      R_g[4,13] := -0.45977530;
      R_g[4,14] := 0.29049909;
      R_g[4,15] := 0.84397930;
      R_g[5,0] := 0.11107527;
      R_g[5,1] := 0.19470578;
      R_g[5,2] := -0.14108169;
      R_g[5,3] := 0.05879988;
      R_g[5,4] := 0.18819207;
      R_g[5,5] := -2.47536159;
      R_g[5,6] := -0.06510852;
      R_g[5,7] := 0.20388806;
      R_g[5,8] := -0.11789436;
      R_g[5,9] := -0.20122005;
      R_g[5,10] := 0.13310707;
      R_g[5,11] := 0.10226060;
      R_g[5,12] := 0.11609720;
      R_g[5,13] := -0.01743704;
      R_g[5,14] := 0.00398547;
      R_g[5,15] := -0.15065657;
      R_g[6,0] := 0.01830370;
      R_g[6,1] := -0.12926060;
      R_g[6,2] := 0.03696303;
      R_g[6,3] := 0.16922043;
      R_g[6,4] := -0.01032830;
      R_g[6,5] := 0.17732817;
      R_g[6,6] := -2.69588876;
      R_g[6,7] := 0.02693873;
      R_g[6,8] := 0.12963313;
      R_g[6,9] := -0.13445157;
      R_g[6,10] := 0.03944382;
      R_g[6,11] := 0.48681569;
      R_g[6,12] := -0.06957243;
      R_g[6,13] := 0.15626159;
      R_g[6,14] := 0.08367650;
      R_g[6,15] := 0.12336652;
      R_g[7,0] := -0.03125253;
      R_g[7,1] := -0.06615835;
      R_g[7,2] := -0.30859804;
      R_g[7,3] := -0.25204793;
      R_g[7,4] := 0.40157086;
      R_g[7,5] := 0.02905789;
      R_g[7,6] := -0.05298730;
      R_g[7,7] := -3.66701341;
      R_g[7,8] := -0.20909342;
      R_g[7,9] := 0.39114916;
      R_g[7,10] := 0.02195679;
      R_g[7,11] := 0.36044669;
      R_g[7,12] := -0.19184318;
      R_g[7,13] := 0.29045779;
      R_g[7,14] := -0.39132181;
      R_g[7,15] := 0.18133201;
      R_g[8,0] := 0.10109203;
      R_g[8,1] := 0.70265359;
      R_g[8,2] := -0.20131305;
      R_g[8,3] := -0.26565599;
      R_g[8,4] := -0.09981477;
      R_g[8,5] := 0.02134162;
      R_g[8,6] := 0.03664974;
      R_g[8,7] := -0.10195713;
      R_g[8,8] := -2.91001201;
      R_g[8,9] := 0.11249696;
      R_g[8,10] := 0.27498955;
      R_g[8,11] := -0.21615753;
      R_g[8,12] := 0.21132010;
      R_g[8,13] := -0.04111291;
      R_g[8,14] := 0.16867815;
      R_g[8,15] := -0.19916441;
      R_g[9,0] := -0.17235202;
      R_g[9,1] := -0.51918679;
      R_g[9,2] := 0.09489006;
      R_g[9,3] := 0.27006283;
      R_g[9,4] := -0.08789669;
      R_g[9,5] := 0.00435399;
      R_g[9,6] := 0.16746791;
      R_g[9,7] := -0.05963518;
      R_g[9,8] := -0.02752298;
      R_g[9,9] := -4.96825457;
      R_g[9,10] := -0.22408967;
      R_g[9,11] := 0.39007574;
      R_g[9,12] := 0.04636907;
      R_g[9,13] := 0.04828465;
      R_g[9,14] := -0.23503923;
      R_g[9,15] := 0.62594104;
      R_g[10,0] := -0.15698923;
      R_g[10,1] := 0.66038901;
      R_g[10,2] := -0.36404622;
      R_g[10,3] := -0.15719211;
      R_g[10,4] := 0.19071013;
      R_g[10,5] := -0.04058476;
      R_g[10,6] := -0.03078617;
      R_g[10,7] := 0.71735823;
      R_g[10,8] := -0.29184514;
      R_g[10,9] := -0.10818060;
      R_g[10,10] := -3.58587956;
      R_g[10,11] := -0.47085500;
      R_g[10,12] := 0.49304882;
      R_g[10,13] := 0.30396828;
      R_g[10,14] := 0.08089786;
      R_g[10,15] := -0.43142110;
      R_g[11,0] := 0.06635704;
      R_g[11,1] := 0.43992752;
      R_g[11,2] := 0.07202107;
      R_g[11,3] := -0.23624249;
      R_g[11,4] := -0.07328893;
      R_g[11,5] := -0.04814436;
      R_g[11,6] := -0.09117863;
      R_g[11,7] := 0.11876864;
      R_g[11,8] := 0.00884132;
      R_g[11,9] := -0.18132856;
      R_g[11,10] := 0.01293289;
      R_g[11,11] := -3.54570603;
      R_g[11,12] := -0.03885806;
      R_g[11,13] := -0.05033415;
      R_g[11,14] := 0.11649126;
      R_g[11,15] := -0.00223985;
      R_g[12,0] := -0.17420630;
      R_g[12,1] := -0.13533008;
      R_g[12,2] := -0.02006780;
      R_g[12,3] := 0.22674133;
      R_g[12,4] := -0.14372772;
      R_g[12,5] := 0.17432602;
      R_g[12,6] := 0.28012389;
      R_g[12,7] := -0.08454837;
      R_g[12,8] := 0.17622249;
      R_g[12,9] := -0.18562099;
      R_g[12,10] := -0.13753660;
      R_g[12,11] := 0.31376547;
      R_g[12,12] := -2.33639669;
      R_g[12,13] := -0.37101883;
      R_g[12,14] := -0.10402304;
      R_g[12,15] := 0.34098265;
      R_g[13,0] := 0.05532536;
      R_g[13,1] := -1.13573086;
      R_g[13,2] := 0.05515465;
      R_g[13,3] := 0.17128730;
      R_g[13,4] := 0.29013124;
      R_g[13,5] := 0.14211339;
      R_g[13,6] := -0.12067565;
      R_g[13,7] := 0.06888673;
      R_g[13,8] := -0.19051172;
      R_g[13,9] := -0.08930715;
      R_g[13,10] := -0.03726633;
      R_g[13,11] := 0.10250945;
      R_g[13,12] := 0.01444966;
      R_g[13,13] := -2.59691453;
      R_g[13,14] := -0.05213837;
      R_g[13,15] := -0.16357523;
      R_g[14,0] := -0.07426858;
      R_g[14,1] := 0.95711172;
      R_g[14,2] := -0.52914786;
      R_g[14,3] := -0.50707346;
      R_g[14,4] := -0.18582524;
      R_g[14,5] := 0.04817829;
      R_g[14,6] := -0.18424018;
      R_g[14,7] := 0.31674099;
      R_g[14,8] := -0.00767360;
      R_g[14,9] := -0.00882705;
      R_g[14,10] := -0.06244185;
      R_g[14,11] := -0.83984315;
      R_g[14,12] := -0.04242671;
      R_g[14,13] := 0.06255507;
      R_g[14,14] := -2.18376112;
      R_g[14,15] := -0.50745595;
      R_g[15,0] := -0.24544616;
      R_g[15,1] := -0.38065434;
      R_g[15,2] := 0.52168375;
      R_g[15,3] := 0.63476181;
      R_g[15,4] := -0.70045185;
      R_g[15,5] := 0.03916581;
      R_g[15,6] := 0.27065009;
      R_g[15,7] := -0.15145577;
      R_g[15,8] := 0.19062088;
      R_g[15,9] := -0.16805187;
      R_g[15,10] := -0.02476993;
      R_g[15,11] := 0.03592181;
      R_g[15,12] := -0.40066659;
      R_g[15,13] := -0.61348122;
      R_g[15,14] := 0.08364772;
      R_g[15,15] := -3.36107063;
      R_o[0,0] := -0.17998135;
      R_o[0,1] := -1.60253966;
      R_o[0,2] := 0.68840933;
      R_o[0,3] := 0.60407180;
      R_o[0,4] := -0.62490994;
      R_o[0,5] := 0.50324053;
      R_o[0,6] := 0.24965659;
      R_o[0,7] := 0.27685815;
      R_o[0,8] := -0.37989971;
      R_o[0,9] := 0.13533561;
      R_o[0,10] := -0.25785661;
      R_o[0,11] := -0.51081169;
      R_o[0,12] := -1.26113296;
      R_o[0,13] := 0.09709056;
      R_o[0,14] := 0.61411685;
      R_o[0,15] := 0.22855295;
      R_o[1,0] := 0.22900739;
      R_o[1,1] := -3.14904022;
      R_o[1,2] := 0.71979213;
      R_o[1,3] := 0.13460559;
      R_o[1,4] := 0.28159738;
      R_o[1,5] := -1.25828946;
      R_o[1,6] := 0.70830607;
      R_o[1,7] := -0.61551344;
      R_o[1,8] := -0.20931304;
      R_o[1,9] := 0.84665543;
      R_o[1,10] := -0.58804363;
      R_o[1,11] := -0.01368906;
      R_o[1,12] := -0.09546302;
      R_o[1,13] := 0.68291515;
      R_o[1,14] := 0.83152312;
      R_o[1,15] := -0.27614936;
      R_o[2,0] := 0.22624512;
      R_o[2,1] := -0.50015140;
      R_o[2,2] := -0.05820123;
      R_o[2,3] := 0.24992104;
      R_o[2,4] := -0.42781389;
      R_o[2,5] := -0.01809851;
      R_o[2,6] := -0.01348706;
      R_o[2,7] := -0.39746183;
      R_o[2,8] := -0.21094593;
      R_o[2,9] := 0.74206448;
      R_o[2,10] := 0.08259194;
      R_o[2,11] := -0.43268228;
      R_o[2,12] := -0.06109180;
      R_o[2,13] := -0.26904088;
      R_o[2,14] := 0.29712129;
      R_o[2,15] := -0.07692748;
      R_o[3,0] := 0.14433832;
      R_o[3,1] := -0.80342203;
      R_o[3,2] := 0.15820050;
      R_o[3,3] := 0.08200698;
      R_o[3,4] := -0.48171204;
      R_o[3,5] := -0.11591465;
      R_o[3,6] := -0.19669321;
      R_o[3,7] := -0.14903167;
      R_o[3,8] := -0.15372486;
      R_o[3,9] := 0.14865009;
      R_o[3,10] := -0.82148689;
      R_o[3,11] := 0.27812725;
      R_o[3,12] := 0.00223510;
      R_o[3,13] := 0.21079217;
      R_o[3,14] := -0.25288963;
      R_o[3,15] := -0.22805665;
      R_o[4,0] := 0.25114408;
      R_o[4,1] := -0.04965499;
      R_o[4,2] := -0.07762759;
      R_o[4,3] := 0.18927185;
      R_o[4,4] := 0.10361283;
      R_o[4,5] := -0.03912014;
      R_o[4,6] := -0.91816306;
      R_o[4,7] := 0.15886311;
      R_o[4,8] := 0.42278275;
      R_o[4,9] := 0.42559728;
      R_o[4,10] := -0.16750900;
      R_o[4,11] := -0.82801008;
      R_o[4,12] := 0.47436076;
      R_o[4,13] := 0.45988649;
      R_o[4,14] := 0.03260082;
      R_o[4,15] := -0.05795699;
      R_o[5,0] := 0.01105135;
      R_o[5,1] := -1.15132201;
      R_o[5,2] := 0.54602605;
      R_o[5,3] := 0.71394539;
      R_o[5,4] := -0.17321546;
      R_o[5,5] := -0.52846497;
      R_o[5,6] := -0.43260244;
      R_o[5,7] := 0.35832340;
      R_o[5,8] := 0.21435645;
      R_o[5,9] := 0.26636124;
      R_o[5,10] := 0.00893501;
      R_o[5,11] := -0.63832158;
      R_o[5,12] := -0.11683670;
      R_o[5,13] := -0.02273753;
      R_o[5,14] := 0.03232908;
      R_o[5,15] := 0.10529289;
      R_o[6,0] := 0.31001085;
      R_o[6,1] := -1.19092143;
      R_o[6,2] := 0.21876206;
      R_o[6,3] := 0.33240157;
      R_o[6,4] := -0.18906151;
      R_o[6,5] := 0.48293993;
      R_o[6,6] := -0.03892522;
      R_o[6,7] := -0.35924369;
      R_o[6,8] := 0.12160594;
      R_o[6,9] := -0.40936342;
      R_o[6,10] := 0.12075932;
      R_o[6,11] := -0.49636525;
      R_o[6,12] := -0.13716739;
      R_o[6,13] := 0.06098676;
      R_o[6,14] := -0.27069107;
      R_o[6,15] := 0.41007137;
      R_o[7,0] := 0.29690558;
      R_o[7,1] := -0.37541282;
      R_o[7,2] := 0.24571100;
      R_o[7,3] := 0.23365253;
      R_o[7,4] := 0.21465455;
      R_o[7,5] := 0.03528690;
      R_o[7,6] := -0.12078243;
      R_o[7,7] := -0.03139850;
      R_o[7,8] := 0.10045099;
      R_o[7,9] := -0.14713535;
      R_o[7,10] := -0.18440804;
      R_o[7,11] := 0.56326222;
      R_o[7,12] := -0.29376999;
      R_o[7,13] := 0.06893768;
      R_o[7,14] := 0.13139424;
      R_o[7,15] := 0.26108429;
      R_o[8,0] := -1.83918154;
      R_o[8,1] := -1.09582520;
      R_o[8,2] := 0.50053239;
      R_o[8,3] := 0.73636478;
      R_o[8,4] := -0.94267857;
      R_o[8,5] := -1.52087641;
      R_o[8,6] := 2.80385971;
      R_o[8,7] := 0.62324148;
      R_o[8,8] := -3.54411769;
      R_o[8,9] := -0.25437289;
      R_o[8,10] := -0.15810332;
      R_o[8,11] := -0.51360112;
      R_o[8,12] := 0.01348928;
      R_o[8,13] := 0.22060399;
      R_o[8,14] := -0.52212816;
      R_o[8,15] := 0.10016742;
      R_o[9,0] := -1.07547414;
      R_o[9,1] := -1.28275371;
      R_o[9,2] := 0.35765028;
      R_o[9,3] := 0.44110700;
      R_o[9,4] := -0.91392058;
      R_o[9,5] := -1.19914532;
      R_o[9,6] := 0.03312799;
      R_o[9,7] := 0.26320797;
      R_o[9,8] := -0.30888504;
      R_o[9,9] := -3.75967288;
      R_o[9,10] := -0.26503733;
      R_o[9,11] := -0.14797226;
      R_o[9,12] := -0.29307473;
      R_o[9,13] := 0.29319406;
      R_o[9,14] := 0.47096246;
      R_o[9,15] := 0.08412670;
      R_o[10,0] := 0.03535339;
      R_o[10,1] := -0.81770265;
      R_o[10,2] := -0.41774553;
      R_o[10,3] := 0.28629521;
      R_o[10,4] := -0.29024190;
      R_o[10,5] := -0.30073890;
      R_o[10,6] := 0.06244223;
      R_o[10,7] := -0.86978775;
      R_o[10,8] := 0.56519794;
      R_o[10,9] := 0.02823679;
      R_o[10,10] := 0.43152261;
      R_o[10,11] := -0.52289534;
      R_o[10,12] := -0.92306936;
      R_o[10,13] := -0.11299136;
      R_o[10,14] := -0.46108496;
      R_o[10,15] := 0.27689543;
      R_o[11,0] := -0.27377477;
      R_o[11,1] := -1.38200986;
      R_o[11,2] := 0.80172545;
      R_o[11,3] := 0.47983712;
      R_o[11,4] := -0.61602306;
      R_o[11,5] := 0.14996068;
      R_o[11,6] := -0.27008256;
      R_o[11,7] := 0.01958398;
      R_o[11,8] := 0.95527297;
      R_o[11,9] := -0.14984407;
      R_o[11,10] := -0.12444744;
      R_o[11,11] := 2.54292870;
      R_o[11,12] := -0.39212865;
      R_o[11,13] := -1.04945409;
      R_o[11,14] := 0.45311722;
      R_o[11,15] := 0.23906973;
      R_o[12,0] := -0.03170222;
      R_o[12,1] := -0.25899503;
      R_o[12,2] := -0.00625280;
      R_o[12,3] := 0.20854484;
      R_o[12,4] := -0.24143498;
      R_o[12,5] := 0.10468624;
      R_o[12,6] := -0.20445421;
      R_o[12,7] := 0.37825984;
      R_o[12,8] := 0.04627231;
      R_o[12,9] := 0.02643433;
      R_o[12,10] := -0.13525262;
      R_o[12,11] := -0.51159739;
      R_o[12,12] := 0.17827436;
      R_o[12,13] := 0.03084075;
      R_o[12,14] := 0.28973144;
      R_o[12,15] := -0.25529897;
      R_o[13,0] := 0.00229840;
      R_o[13,1] := -1.61626279;
      R_o[13,2] := 0.40775979;
      R_o[13,3] := 0.59826922;
      R_o[13,4] := -0.21434167;
      R_o[13,5] := -0.15114538;
      R_o[13,6] := -0.73304671;
      R_o[13,7] := -0.11104193;
      R_o[13,8] := -0.43963873;
      R_o[13,9] := 0.18838404;
      R_o[13,10] := 0.39571330;
      R_o[13,11] := -1.05748773;
      R_o[13,12] := -0.32323301;
      R_o[13,13] := 1.01370287;
      R_o[13,14] := 0.21895173;
      R_o[13,15] := 0.80038011;
      R_o[14,0] := -0.07648548;
      R_o[14,1] := -1.30468404;
      R_o[14,2] := 0.58321625;
      R_o[14,3] := 0.72309285;
      R_o[14,4] := 0.12278607;
      R_o[14,5] := 0.20592272;
      R_o[14,6] := -1.31852913;
      R_o[14,7] := -0.26429388;
      R_o[14,8] := 0.67733824;
      R_o[14,9] := 0.28490099;
      R_o[14,10] := 0.50044572;
      R_o[14,11] := 1.13938892;
      R_o[14,12] := -0.62636727;
      R_o[14,13] := -0.64233524;
      R_o[14,14] := 2.21524429;
      R_o[14,15] := 0.10953581;
      R_o[15,0] := -0.61134338;
      R_o[15,1] := -1.14686418;
      R_o[15,2] := 0.91901773;
      R_o[15,3] := 0.59483540;
      R_o[15,4] := -1.43020630;
      R_o[15,5] := -0.02133927;
      R_o[15,6] := 0.24188809;
      R_o[15,7] := -0.50801885;
      R_o[15,8] := 0.25780970;
      R_o[15,9] := 0.13150303;
      R_o[15,10] := 0.06579445;
      R_o[15,11] := 0.21622118;
      R_o[15,12] := -0.23762867;
      R_o[15,13] := -0.99601251;
      R_o[15,14] := 0.53441352;
      R_o[15,15] := 2.04913473;
      B_i[0] := 2.13055468;
      B_i[1] := -0.28939855;
      B_i[2] := 2.50660825;
      B_i[3] := -0.09900541;
      B_i[4] := 0.92722613;
      B_i[5] := -0.24022682;
      B_i[6] := 0.01314271;
      B_i[7] := -0.16002662;
      B_i[8] := -0.13514934;
      B_i[9] := -0.66461527;
      B_i[10] := -0.39439538;
      B_i[11] := -0.72713459;
      B_i[12] := 2.69549060;
      B_i[13] := 0.10082641;
      B_i[14] := 0.18705003;
      B_i[15] := -0.52215415;
      B_f[0] := 1.71853232;
      B_f[1] := 0.52807707;
      B_f[2] := -0.91032523;
      B_f[3] := -0.51656717;
      B_f[4] := 3.52749252;
      B_f[5] := 2.54868436;
      B_f[6] := 2.06901407;
      B_f[7] := 4.24917698;
      B_f[8] := 2.06338930;
      B_f[9] := 2.86993122;
      B_f[10] := 3.17252159;
      B_f[11] := 1.42340124;
      B_f[12] := 4.81506538;
      B_f[13] := 1.14250445;
      B_f[14] := 0.49386898;
      B_f[15] := 2.75026822;
      B_g[0] := -0.07227773;
      B_g[1] := -0.66488314;
      B_g[2] := 0.70045793;
      B_g[3] := 0.98024452;
      B_g[4] := -0.46857694;
      B_g[5] := 0.02956967;
      B_g[6] := 0.27909416;
      B_g[7] := -0.22752739;
      B_g[8] := -0.10114017;
      B_g[9] := -0.10326473;
      B_g[10] := 0.06763726;
      B_g[11] := 0.14730735;
      B_g[12] := -0.17682402;
      B_g[13] := -0.28040373;
      B_g[14] := 0.69763172;
      B_g[15] := -0.60094702;
      B_o[0] := 3.63638949;
      B_o[1] := 3.95470619;
      B_o[2] := 2.86919069;
      B_o[3] := 2.67019081;
      B_o[4] := 2.45756173;
      B_o[5] := 2.80873203;
      B_o[6] := 2.80962849;
      B_o[7] := 1.47691143;
      B_o[8] := 4.80254173;
      B_o[9] := 3.77295828;
      B_o[10] := 3.93514633;
      B_o[11] := 3.18298674;
      B_o[12] := 1.06958044;
      B_o[13] := 3.72094917;
      B_o[14] := 2.60961676;
      B_o[15] := 3.24567151;
      FC_W[0,0] := -0.82467866;
      FC_W[0,1] := 0.23118977;
      FC_W[0,2] := -0.56444192;
      FC_W[0,3] := -0.32562086;
      FC_W[0,4] := 0.93298566;
      FC_W[0,5] := -1.32120907;
      FC_W[0,6] := -0.26805392;
      FC_W[0,7] := -0.71825963;
      FC_W[0,8] := -1.19989681;
      FC_W[0,9] := -2.48990393;
      FC_W[0,10] := 0.54710686;
      FC_W[0,11] := -1.50483215;
      FC_W[0,12] := -0.24574320;
      FC_W[0,13] := 1.17454255;
      FC_W[0,14] := 0.51390719;
      FC_W[0,15] := 1.51483810;
      FC_W[1,0] := 1.04243851;
      FC_W[1,1] := 1.69587207;
      FC_W[1,2] := 1.49340200;
      FC_W[1,3] := -1.27457929;
      FC_W[1,4] := -0.06108139;
      FC_W[1,5] := 0.15937902;
      FC_W[1,6] := -0.56430584;
      FC_W[1,7] := -1.76767778;
      FC_W[1,8] := 0.98803681;
      FC_W[1,9] := -0.39248836;
      FC_W[1,10] := 1.23283052;
      FC_W[1,11] := 2.07260656;
      FC_W[1,12] := -1.40971696;
      FC_W[1,13] := -1.29698300;
      FC_W[1,14] := 2.06386137;
      FC_W[1,15] := -0.25542155;
      FC_W[2,0] := -0.85026604;
      FC_W[2,1] := 0.35434592;
      FC_W[2,2] := -0.44842285;
      FC_W[2,3] := -0.44237766;
      FC_W[2,4] := 0.85990745;
      FC_W[2,5] := -1.32394731;
      FC_W[2,6] := -0.31900164;
      FC_W[2,7] := -0.75662905;
      FC_W[2,8] := -1.19999981;
      FC_W[2,9] := -2.58493805;
      FC_W[2,10] := 0.55032092;
      FC_W[2,11] := -1.63180840;
      FC_W[2,12] := -0.31313592;
      FC_W[2,13] := 1.21769071;
      FC_W[2,14] := 0.62405908;
      FC_W[2,15] := 1.54905689;
      FC_W[3,0] := 0.17799814;
      FC_W[3,1] := 0.31846881;
      FC_W[3,2] := 0.10473058;
      FC_W[3,3] := -0.13281064;
      FC_W[3,4] := -0.17808376;
      FC_W[3,5] := 1.50857568;
      FC_W[3,6] := 0.46525395;
      FC_W[3,7] := 0.05502938;
      FC_W[3,8] := -0.57212090;
      FC_W[3,9] := -2.09590507;
      FC_W[3,10] := -0.40869591;
      FC_W[3,11] := 0.00603901;
      FC_W[3,12] := 0.39652750;
      FC_W[3,13] := 0.60246611;
      FC_W[3,14] := -1.03614700;
      FC_W[3,15] := 0.55060035;
      FC_W[4,0] := 1.10157812;
      FC_W[4,1] := -0.82706159;
      FC_W[4,2] := 0.62553823;
      FC_W[4,3] := -0.65783793;
      FC_W[4,4] := -0.42305151;
      FC_W[4,5] := -0.49417713;
      FC_W[4,6] := 0.27170289;
      FC_W[4,7] := 0.77937496;
      FC_W[4,8] := 1.34962928;
      FC_W[4,9] := -0.56700414;
      FC_W[4,10] := -2.24635792;
      FC_W[4,11] := -0.41298652;
      FC_W[4,12] := -0.51241404;
      FC_W[4,13] := -1.14208841;
      FC_W[4,14] := -0.00704930;
      FC_W[4,15] := 1.58584416;
      FC_W[5,0] := 0.04869050;
      FC_W[5,1] := -2.49297285;
      FC_W[5,2] := -0.44874841;
      FC_W[5,3] := 0.17483039;
      FC_W[5,4] := 0.22983202;
      FC_W[5,5] := -2.60724688;
      FC_W[5,6] := -0.43566737;
      FC_W[5,7] := 2.92718530;
      FC_W[5,8] := 3.13831282;
      FC_W[5,9] := -3.70684314;
      FC_W[5,10] := -0.49225014;
      FC_W[5,11] := 0.98027021;
      FC_W[5,12] := 0.85220718;
      FC_W[5,13] := -0.35435688;
      FC_W[5,14] := -0.21338330;
      FC_W[5,15] := -3.31668758;
      FC_W[6,0] := 0.58065802;
      FC_W[6,1] := 0.58166015;
      FC_W[6,2] := 0.29509109;
      FC_W[6,3] := 1.24706650;
      FC_W[6,4] := 0.32439369;
      FC_W[6,5] := 0.15459089;
      FC_W[6,6] := 0.11035646;
      FC_W[6,7] := 2.14783597;
      FC_W[6,8] := 0.13601644;
      FC_W[6,9] := -1.02714729;
      FC_W[6,10] := 0.23564745;
      FC_W[6,11] := 0.42390209;
      FC_W[6,12] := -0.84225869;
      FC_W[6,13] := 0.07522085;
      FC_W[6,14] := -0.27497068;
      FC_W[6,15] := 0.15566382;
      FC_W[7,0] := 0.18631160;
      FC_W[7,1] := 0.25749409;
      FC_W[7,2] := 0.05877232;
      FC_W[7,3] := -0.08437430;
      FC_W[7,4] := -0.14088097;
      FC_W[7,5] := 1.50284660;
      FC_W[7,6] := 0.48287323;
      FC_W[7,7] := 0.08982904;
      FC_W[7,8] := -0.56427842;
      FC_W[7,9] := -2.04194164;
      FC_W[7,10] := -0.43468520;
      FC_W[7,11] := 0.05047191;
      FC_W[7,12] := 0.41730252;
      FC_W[7,13] := 0.59546208;
      FC_W[7,14] := -1.09572983;
      FC_W[7,15] := 0.53943986;
      FC_W[8,0] := 0.17352782;
      FC_W[8,1] := 0.42593235;
      FC_W[8,2] := 0.11490290;
      FC_W[8,3] := -0.25036201;
      FC_W[8,4] := -0.17699352;
      FC_W[8,5] := 1.51737905;
      FC_W[8,6] := 0.45302224;
      FC_W[8,7] := 0.02927133;
      FC_W[8,8] := -0.58808583;
      FC_W[8,9] := -2.18285322;
      FC_W[8,10] := -0.37657666;
      FC_W[8,11] := -0.04062983;
      FC_W[8,12] := 0.41792968;
      FC_W[8,13] := 0.55557293;
      FC_W[8,14] := -0.95937282;
      FC_W[8,15] := 0.55914086;
      FC_W[9,0] := 0.17505446;
      FC_W[9,1] := 0.28600723;
      FC_W[9,2] := 0.07933394;
      FC_W[9,3] := -0.12126631;
      FC_W[9,4] := -0.15457296;
      FC_W[9,5] := 1.50301993;
      FC_W[9,6] := 0.47192392;
      FC_W[9,7] := 0.06274927;
      FC_W[9,8] := -0.56979150;
      FC_W[9,9] := -2.07217526;
      FC_W[9,10] := -0.41918421;
      FC_W[9,11] := 0.03827762;
      FC_W[9,12] := 0.41007796;
      FC_W[9,13] := 0.60690254;
      FC_W[9,14] := -1.06829190;
      FC_W[9,15] := 0.53677040;
      FC_W[10,0] := -0.25367916;
      FC_W[10,1] := -0.32994914;
      FC_W[10,2] := -0.15668485;
      FC_W[10,3] := -1.45790470;
      FC_W[10,4] := -0.16369641;
      FC_W[10,5] := 0.29133776;
      FC_W[10,6] := 0.14205573;
      FC_W[10,7] := -0.87707573;
      FC_W[10,8] := 0.42122248;
      FC_W[10,9] := -3.06178594;
      FC_W[10,10] := -0.44065821;
      FC_W[10,11] := 0.50379735;
      FC_W[10,12] := 1.11131394;
      FC_W[10,13] := 0.31328326;
      FC_W[10,14] := -0.66578966;
      FC_W[10,15] := -0.78003192;
      FC_W[11,0] := 0.13824168;
      FC_W[11,1] := 0.30625078;
      FC_W[11,2] := 0.69278711;
      FC_W[11,3] := -0.47781393;
      FC_W[11,4] := -0.95308739;
      FC_W[11,5] := 0.04460392;
      FC_W[11,6] := 0.38477588;
      FC_W[11,7] := 0.07937323;
      FC_W[11,8] := -1.41032720;
      FC_W[11,9] := -0.44885933;
      FC_W[11,10] := -0.81729096;
      FC_W[11,11] := 0.41849750;
      FC_W[11,12] := -1.37481093;
      FC_W[11,13] := -0.12758188;
      FC_W[11,14] := -0.37933919;
      FC_W[11,15] := -0.96544886;
      FC_W[12,0] := -0.33354285;
      FC_W[12,1] := 0.31888646;
      FC_W[12,2] := 1.15725291;
      FC_W[12,3] := -0.57309943;
      FC_W[12,4] := -0.63576299;
      FC_W[12,5] := 0.31176066;
      FC_W[12,6] := 0.16692483;
      FC_W[12,7] := 0.08488149;
      FC_W[12,8] := -0.91559130;
      FC_W[12,9] := -0.37182277;
      FC_W[12,10] := -0.86818475;
      FC_W[12,11] := 0.33183327;
      FC_W[12,12] := -1.33442044;
      FC_W[12,13] := 0.02328874;
      FC_W[12,14] := -0.47359598;
      FC_W[12,15] := -0.85911077;
      FC_W[13,0] := 0.34582901;
      FC_W[13,1] := -1.24973571;
      FC_W[13,2] := 0.09938692;
      FC_W[13,3] := 0.27242026;
      FC_W[13,4] := 2.86735916;
      FC_W[13,5] := -1.29841161;
      FC_W[13,6] := -0.55971164;
      FC_W[13,7] := -1.16741526;
      FC_W[13,8] := -0.10935560;
      FC_W[13,9] := 0.36287791;
      FC_W[13,10] := 0.64087117;
      FC_W[13,11] := 4.35670900;
      FC_W[13,12] := -0.46027356;
      FC_W[13,13] := 1.15009689;
      FC_W[13,14] := 0.52797776;
      FC_W[13,15] := -0.36370721;
      FC_W[14,0] := -3.52245569;
      FC_W[14,1] := -1.56672299;
      FC_W[14,2] := -3.15010047;
      FC_W[14,3] := -0.65020859;
      FC_W[14,4] := -0.49099338;
      FC_W[14,5] := 3.08911586;
      FC_W[14,6] := 1.92608213;
      FC_W[14,7] := 0.08825259;
      FC_W[14,8] := 0.54131156;
      FC_W[14,9] := -0.49000683;
      FC_W[14,10] := -1.64109290;
      FC_W[14,11] := 0.88520831;
      FC_W[14,12] := -1.96192515;
      FC_W[14,13] := -0.16477479;
      FC_W[14,14] := 2.96418428;
      FC_W[14,15] := 0.30263656;
      FC_W[15,0] := 0.74186748;
      FC_W[15,1] := 0.62531567;
      FC_W[15,2] := 0.26485214;
      FC_W[15,3] := -0.18005861;
      FC_W[15,4] := -1.44341528;
      FC_W[15,5] := -0.49698487;
      FC_W[15,6] := 0.51499581;
      FC_W[15,7] := 0.11231317;
      FC_W[15,8] := -1.84129775;
      FC_W[15,9] := -0.48331323;
      FC_W[15,10] := -0.82623559;
      FC_W[15,11] := 0.57879627;
      FC_W[15,12] := -1.45617056;
      FC_W[15,13] := 0.34439510;
      FC_W[15,14] := -0.02835772;
      FC_W[15,15] := -0.95853078;
      FC_W[16,0] := -0.10502820;
      FC_W[16,1] := 2.86326361;
      FC_W[16,2] := 0.41696814;
      FC_W[16,3] := 0.68216890;
      FC_W[16,4] := -1.25698853;
      FC_W[16,5] := -1.68472195;
      FC_W[16,6] := 2.72576451;
      FC_W[16,7] := -0.13771258;
      FC_W[16,8] := 2.13751483;
      FC_W[16,9] := -0.05118477;
      FC_W[16,10] := -0.69813430;
      FC_W[16,11] := 0.59181178;
      FC_W[16,12] := -0.59705693;
      FC_W[16,13] := 5.95551205;
      FC_W[16,14] := 0.87344640;
      FC_W[16,15] := 1.47654462;
      FC_W[17,0] := -3.72690654;
      FC_W[17,1] := -0.34288198;
      FC_W[17,2] := 3.20892954;
      FC_W[17,3] := -1.09288120;
      FC_W[17,4] := 2.75555611;
      FC_W[17,5] := 1.44968975;
      FC_W[17,6] := 0.08937956;
      FC_W[17,7] := -0.05114520;
      FC_W[17,8] := 3.77698874;
      FC_W[17,9] := 0.68791342;
      FC_W[17,10] := -0.32791337;
      FC_W[17,11] := -1.15987170;
      FC_W[17,12] := 0.12185520;
      FC_W[17,13] := 0.77343524;
      FC_W[17,14] := -0.91215330;
      FC_W[17,15] := 0.44880545;
      FC_W[18,0] := -0.36295000;
      FC_W[18,1] := 0.59718996;
      FC_W[18,2] := -2.02808356;
      FC_W[18,3] := 0.21908940;
      FC_W[18,4] := -0.35514835;
      FC_W[18,5] := -0.16581751;
      FC_W[18,6] := 0.32898539;
      FC_W[18,7] := -1.00391436;
      FC_W[18,8] := 2.15731025;
      FC_W[18,9] := -0.97810787;
      FC_W[18,10] := 0.30121070;
      FC_W[18,11] := -0.79974371;
      FC_W[18,12] := -4.20807362;
      FC_W[18,13] := -1.48771405;
      FC_W[18,14] := -5.74529266;
      FC_W[18,15] := -0.61625999;
      FC_W[19,0] := -0.42781910;
      FC_W[19,1] := 0.01137099;
      FC_W[19,2] := 1.65118229;
      FC_W[19,3] := -0.67069191;
      FC_W[19,4] := -0.41222230;
      FC_W[19,5] := 0.51861578;
      FC_W[19,6] := -0.32404739;
      FC_W[19,7] := 0.37804386;
      FC_W[19,8] := -1.31013584;
      FC_W[19,9] := -0.10698038;
      FC_W[19,10] := -0.96316320;
      FC_W[19,11] := 0.46424603;
      FC_W[19,12] := -0.41702995;
      FC_W[19,13] := -0.00965757;
      FC_W[19,14] := 0.69454628;
      FC_W[19,15] := -0.74284571;
      FC_W[20,0] := -0.83391452;
      FC_W[20,1] := -1.79579413;
      FC_W[20,2] := -0.25979164;
      FC_W[20,3] := -1.17057109;
      FC_W[20,4] := -0.70292395;
      FC_W[20,5] := -0.29942927;
      FC_W[20,6] := 0.19507834;
      FC_W[20,7] := -1.58461428;
      FC_W[20,8] := 0.30485892;
      FC_W[20,9] := 1.04576087;
      FC_W[20,10] := -0.16007894;
      FC_W[20,11] := 0.69425857;
      FC_W[20,12] := 0.83975720;
      FC_W[20,13] := -0.30882624;
      FC_W[20,14] := -0.55371881;
      FC_W[20,15] := 0.27732018;
      FC_W[21,0] := -2.10582590;
      FC_W[21,1] := 1.55697012;
      FC_W[21,2] := -0.07022452;
      FC_W[21,3] := 1.33484554;
      FC_W[21,4] := -0.96722597;
      FC_W[21,5] := -0.44053811;
      FC_W[21,6] := 0.60700059;
      FC_W[21,7] := 0.51479501;
      FC_W[21,8] := -1.00228095;
      FC_W[21,9] := -0.81924778;
      FC_W[21,10] := 0.73371696;
      FC_W[21,11] := 0.43934014;
      FC_W[21,12] := 0.41138521;
      FC_W[21,13] := -1.01041663;
      FC_W[21,14] := -0.61670274;
      FC_W[21,15] := 1.38253033;
      FC_W[22,0] := -0.00039924;
      FC_W[22,1] := -1.84598529;
      FC_W[22,2] := 1.43738365;
      FC_W[22,3] := 2.26899028;
      FC_W[22,4] := -0.75990319;
      FC_W[22,5] := 0.37804359;
      FC_W[22,6] := 0.13571464;
      FC_W[22,7] := -0.38089994;
      FC_W[22,8] := 0.59762645;
      FC_W[22,9] := -0.20303242;
      FC_W[22,10] := 0.36337435;
      FC_W[22,11] := 0.81648386;
      FC_W[22,12] := -0.67675233;
      FC_W[22,13] := -0.57171708;
      FC_W[22,14] := 1.22118664;
      FC_W[22,15] := 1.41899049;
      FC_W[23,0] := 0.79800993;
      FC_W[23,1] := -1.77577627;
      FC_W[23,2] := -0.19995016;
      FC_W[23,3] := 0.62975299;
      FC_W[23,4] := 2.48560238;
      FC_W[23,5] := -0.23069511;
      FC_W[23,6] := -0.37795240;
      FC_W[23,7] := -1.11393869;
      FC_W[23,8] := -0.44865733;
      FC_W[23,9] := 0.19626084;
      FC_W[23,10] := 0.59841198;
      FC_W[23,11] := 4.09683037;
      FC_W[23,12] := -0.07720599;
      FC_W[23,13] := 1.75815403;
      FC_W[23,14] := -0.06996297;
      FC_W[23,15] := -0.57559246;
      FC_W[24,0] := -0.02219526;
      FC_W[24,1] := -1.82730865;
      FC_W[24,2] := 1.34180808;
      FC_W[24,3] := 2.47471619;
      FC_W[24,4] := -0.67823833;
      FC_W[24,5] := 0.33719406;
      FC_W[24,6] := 0.16103593;
      FC_W[24,7] := -0.34587914;
      FC_W[24,8] := 0.66295600;
      FC_W[24,9] := -0.14361435;
      FC_W[24,10] := 0.21711408;
      FC_W[24,11] := 0.88477075;
      FC_W[24,12] := -0.77588159;
      FC_W[24,13] := -0.62945527;
      FC_W[24,14] := 0.98504752;
      FC_W[24,15] := 1.34222090;
      FC_W[25,0] := -0.02232726;
      FC_W[25,1] := -1.82818913;
      FC_W[25,2] := 1.34063292;
      FC_W[25,3] := 2.47560835;
      FC_W[25,4] := -0.67833096;
      FC_W[25,5] := 0.33786187;
      FC_W[25,6] := 0.16134858;
      FC_W[25,7] := -0.34436277;
      FC_W[25,8] := 0.66250080;
      FC_W[25,9] := -0.14165786;
      FC_W[25,10] := 0.21584821;
      FC_W[25,11] := 0.88110185;
      FC_W[25,12] := -0.77455860;
      FC_W[25,13] := -0.62910509;
      FC_W[25,14] := 0.98521149;
      FC_W[25,15] := 1.34052444;
      FC_W[26,0] := 1.53153145;
      FC_W[26,1] := -2.05696177;
      FC_W[26,2] := 1.49585950;
      FC_W[26,3] := 0.53426719;
      FC_W[26,4] := 0.46861684;
      FC_W[26,5] := 0.42360222;
      FC_W[26,6] := -0.40656611;
      FC_W[26,7] := -0.34250882;
      FC_W[26,8] := 0.66723526;
      FC_W[26,9] := 0.09229235;
      FC_W[26,10] := -0.06958210;
      FC_W[26,11] := 1.07581246;
      FC_W[26,12] := -0.26606715;
      FC_W[26,13] := 0.61396676;
      FC_W[26,14] := 2.22299767;
      FC_W[26,15] := 0.28380346;
      FC_W[27,0] := -2.24775004;
      FC_W[27,1] := 2.06835508;
      FC_W[27,2] := -0.38080394;
      FC_W[27,3] := 1.01407099;
      FC_W[27,4] := -0.53518450;
      FC_W[27,5] := -0.83131099;
      FC_W[27,6] := 0.66271538;
      FC_W[27,7] := 0.55433625;
      FC_W[27,8] := -1.20186865;
      FC_W[27,9] := -0.79666340;
      FC_W[27,10] := 0.11673751;
      FC_W[27,11] := 0.96070296;
      FC_W[27,12] := 0.87735772;
      FC_W[27,13] := -1.02235091;
      FC_W[27,14] := -0.90932822;
      FC_W[27,15] := 1.24615335;
      FC_W[28,0] := 1.64309812;
      FC_W[28,1] := 0.52149487;
      FC_W[28,2] := 0.80122745;
      FC_W[28,3] := -0.94465780;
      FC_W[28,4] := 0.76917243;
      FC_W[28,5] := -0.94039547;
      FC_W[28,6] := 0.09860569;
      FC_W[28,7] := 1.80428100;
      FC_W[28,8] := 0.30603549;
      FC_W[28,9] := -1.46009111;
      FC_W[28,10] := -1.88728368;
      FC_W[28,11] := 0.87113154;
      FC_W[28,12] := -0.68288696;
      FC_W[28,13] := -0.53775567;
      FC_W[28,14] := 0.81191713;
      FC_W[28,15] := 1.44850564;
      FC_W[29,0] := 0.17561096;
      FC_W[29,1] := 1.04836190;
      FC_W[29,2] := -1.48314321;
      FC_W[29,3] := -1.15159464;
      FC_W[29,4] := 0.95492810;
      FC_W[29,5] := -0.25582403;
      FC_W[29,6] := -0.11323502;
      FC_W[29,7] := 0.75867248;
      FC_W[29,8] := -0.46388596;
      FC_W[29,9] := 0.88885117;
      FC_W[29,10] := -0.88432306;
      FC_W[29,11] := -1.05321443;
      FC_W[29,12] := 0.83339536;
      FC_W[29,13] := 0.75229061;
      FC_W[29,14] := -1.16928649;
      FC_W[29,15] := -1.77717257;
      FC_W[30,0] := 0.00225888;
      FC_W[30,1] := -1.84779334;
      FC_W[30,2] := 1.43843913;
      FC_W[30,3] := 2.26375580;
      FC_W[30,4] := -0.76323915;
      FC_W[30,5] := 0.37884009;
      FC_W[30,6] := 0.13441588;
      FC_W[30,7] := -0.38262546;
      FC_W[30,8] := 0.59856516;
      FC_W[30,9] := -0.20446825;
      FC_W[30,10] := 0.36636823;
      FC_W[30,11] := 0.81112093;
      FC_W[30,12] := -0.67545432;
      FC_W[30,13] := -0.57015026;
      FC_W[30,14] := 1.22726870;
      FC_W[30,15] := 1.41847301;
      FC_W[31,0] := 0.02364270;
      FC_W[31,1] := -1.86203098;
      FC_W[31,2] := 1.46046090;
      FC_W[31,3] := 2.18734074;
      FC_W[31,4] := -0.80845261;
      FC_W[31,5] := 0.41171446;
      FC_W[31,6] := 0.12035200;
      FC_W[31,7] := -0.37572986;
      FC_W[31,8] := 0.57835883;
      FC_W[31,9] := -0.21611637;
      FC_W[31,10] := 0.41468546;
      FC_W[31,11] := 0.72163451;
      FC_W[31,12] := -0.67383784;
      FC_W[31,13] := -0.54498684;
      FC_W[31,14] := 1.29721439;
      FC_W[31,15] := 1.43683994;
      FC_W[32,0] := -0.09428574;
      FC_W[32,1] := -1.68160450;
      FC_W[32,2] := 1.46070540;
      FC_W[32,3] := 2.17403126;
      FC_W[32,4] := -0.76823556;
      FC_W[32,5] := 0.28872356;
      FC_W[32,6] := 0.17703834;
      FC_W[32,7] := -0.35479575;
      FC_W[32,8] := 0.55185831;
      FC_W[32,9] := -0.32400092;
      FC_W[32,10] := 0.35775110;
      FC_W[32,11] := 1.04181564;
      FC_W[32,12] := -0.61921388;
      FC_W[32,13] := -0.68142074;
      FC_W[32,14] := 1.20282924;
      FC_W[32,15] := 1.55295825;
      FC_W[33,0] := -0.11205512;
      FC_W[33,1] := -1.56396496;
      FC_W[33,2] := 1.58497036;
      FC_W[33,3] := 1.87984467;
      FC_W[33,4] := -0.91584122;
      FC_W[33,5] := 0.29638132;
      FC_W[33,6] := 0.17020327;
      FC_W[33,7] := -0.36170369;
      FC_W[33,8] := 0.48853421;
      FC_W[33,9] := -0.47568771;
      FC_W[33,10] := 0.50960517;
      FC_W[33,11] := 0.97275561;
      FC_W[33,12] := -0.53712690;
      FC_W[33,13] := -0.71276188;
      FC_W[33,14] := 1.42409050;
      FC_W[33,15] := 1.71336114;
      FC_W[34,0] := -0.07540017;
      FC_W[34,1] := -1.63697076;
      FC_W[34,2] := 1.53251398;
      FC_W[34,3] := 1.96561730;
      FC_W[34,4] := -0.90749109;
      FC_W[34,5] := 0.33922446;
      FC_W[34,6] := 0.15605466;
      FC_W[34,7] := -0.40329400;
      FC_W[34,8] := 0.53582394;
      FC_W[34,9] := -0.42826504;
      FC_W[34,10] := 0.49411091;
      FC_W[34,11] := 0.84230876;
      FC_W[34,12] := -0.63152224;
      FC_W[34,13] := -0.68104994;
      FC_W[34,14] := 1.34473622;
      FC_W[34,15] := 1.63427615;
      FC_W[35,0] := -0.11846476;
      FC_W[35,1] := -1.67676830;
      FC_W[35,2] := 1.34689760;
      FC_W[35,3] := 2.27766538;
      FC_W[35,4] := -0.63664418;
      FC_W[35,5] := 0.23257758;
      FC_W[35,6] := 0.19841929;
      FC_W[35,7] := -0.36411083;
      FC_W[35,8] := 0.56639081;
      FC_W[35,9] := -0.27044037;
      FC_W[35,10] := 0.27492777;
      FC_W[35,11] := 1.23082864;
      FC_W[35,12] := -0.66170263;
      FC_W[35,13] := -0.67382199;
      FC_W[35,14] := 0.98240697;
      FC_W[35,15] := 1.46826613;
      FC_W[36,0] := -0.07254883;
      FC_W[36,1] := 0.45705366;
      FC_W[36,2] := -0.04096549;
      FC_W[36,3] := 5.95912123;
      FC_W[36,4] := 1.24097335;
      FC_W[36,5] := -0.44737113;
      FC_W[36,6] := 0.09126619;
      FC_W[36,7] := -0.22732373;
      FC_W[36,8] := 0.30773881;
      FC_W[36,9] := 0.21318978;
      FC_W[36,10] := -3.30295229;
      FC_W[36,11] := -0.82223618;
      FC_W[36,12] := -0.09485824;
      FC_W[36,13] := -0.37901035;
      FC_W[36,14] := 0.27817079;
      FC_W[36,15] := -1.09995174;
      FC_W[37,0] := -0.12263552;
      FC_W[37,1] := -1.65574646;
      FC_W[37,2] := 1.31708717;
      FC_W[37,3] := 2.32719302;
      FC_W[37,4] := -0.58871067;
      FC_W[37,5] := 0.21447594;
      FC_W[37,6] := 0.20136184;
      FC_W[37,7] := -0.36005378;
      FC_W[37,8] := 0.56343257;
      FC_W[37,9] := -0.25685868;
      FC_W[37,10] := 0.24374108;
      FC_W[37,11] := 1.28425896;
      FC_W[37,12] := -0.67143738;
      FC_W[37,13] := -0.66641200;
      FC_W[37,14] := 0.92938018;
      FC_W[37,15] := 1.43421566;
      FC_W[38,0] := 0.15314442;
      FC_W[38,1] := 1.63174999;
      FC_W[38,2] := 0.27058762;
      FC_W[38,3] := 0.59943092;
      FC_W[38,4] := -1.74474192;
      FC_W[38,5] := 0.36229685;
      FC_W[38,6] := -5.28263807;
      FC_W[38,7] := 0.33247045;
      FC_W[38,8] := 1.36935079;
      FC_W[38,9] := -0.03816394;
      FC_W[38,10] := -0.68717140;
      FC_W[38,11] := 1.10767031;
      FC_W[38,12] := 0.38817576;
      FC_W[38,13] := 2.73561430;
      FC_W[38,14] := -0.64182931;
      FC_W[38,15] := 2.30720973;
      FC_W[39,0] := -1.88073039;
      FC_W[39,1] := -0.19889264;
      FC_W[39,2] := -1.61357796;
      FC_W[39,3] := 0.00423837;
      FC_W[39,4] := -1.19068766;
      FC_W[39,5] := 2.23228359;
      FC_W[39,6] := -2.08800292;
      FC_W[39,7] := 0.27871919;
      FC_W[39,8] := 1.03275037;
      FC_W[39,9] := -0.31836623;
      FC_W[39,10] := -1.23357213;
      FC_W[39,11] := 0.90982759;
      FC_W[39,12] := -0.73010570;
      FC_W[39,13] := 0.99842566;
      FC_W[39,14] := 1.28712189;
      FC_W[39,15] := 1.49403679;
      FC_B[0] := 0.28719911;
      FC_B[1] := -0.08914877;
      FC_B[2] := 0.27641785;
      FC_B[3] := 0.03852136;
      FC_B[4] := -0.43950242;
      FC_B[5] := 0.24735703;
      FC_B[6] := 0.20127358;
      FC_B[7] := 0.04361544;
      FC_B[8] := 0.07538859;
      FC_B[9] := 0.04495329;
      FC_B[10] := 0.17734325;
      FC_B[11] := -0.63346195;
      FC_B[12] := -0.60759270;
      FC_B[13] := -0.20135863;
      FC_B[14] := 0.53291798;
      FC_B[15] := -0.66306138;
      FC_B[16] := -0.00012068;
      FC_B[17] := 0.09845824;
      FC_B[18] := 1.29676962;
      FC_B[19] := -0.82631814;
      FC_B[20] := -0.47077200;
      FC_B[21] := 0.13384067;
      FC_B[22] := -1.45924211;
      FC_B[23] := -0.31001040;
      FC_B[24] := -1.42507160;
      FC_B[25] := -1.42476630;
      FC_B[26] := -1.19584513;
      FC_B[27] := 0.42283630;
      FC_B[28] := -0.03980854;
      FC_B[29] := 1.16662824;
      FC_B[30] := -1.46038556;
      FC_B[31] := -1.46993387;
      FC_B[32] := -1.42415285;
      FC_B[33] := -1.42881656;
      FC_B[34] := -1.42596591;
      FC_B[35] := -1.37361383;
      FC_B[36] := -0.70964396;
      FC_B[37] := -1.35748100;
      FC_B[38] := 0.86545926;
      FC_B[39] := 0.78649092;

END_DATA_BLOCK
